{attribute 'qualified_only'}
{attribute 'strict'}
{attribute 'to_string'}
TYPE E_PolarIIChamberRotateDirection :
(
	Unknown := 0,
	CW := 1,
	CCW := 2
) UINT;
END_TYPE

(* stored: Version 1.1.0.1, ProductVersion 3.1.4026.18
   DUT E_PolarIIChamberRotateDirection: Id {14000000-0000-0000-0000-000000000004} *)
